TYPE "FRK_SequenceRow"
VERSION : 0.1
   STRUCT
      StepNo : DInt;
      Visited : Bool;
      LastDuration : Time;
   END_STRUCT;

END_TYPE

